Fanuc KAREL source: KT00170.KL

PROGRAM KT00170
%NOLOCKGROUP
VAR
  R1: REAL
  I2: INTEGER
  OUT: REAL
BEGIN
  R1 = 2.0
    I2 = 3
  OUT = R1 MOD I2
END KT00170
